FUNCTION_BLOCK Processing2CAT (* CAT Function Block Type *)
  (* Standard: 61499-2 *)
  (* Version 0.0, 7/7/2026, template *)
  PACKAGE Main;
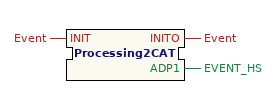
  EVENT_INPUT
    INIT; (* Initialization Request *)
  END_EVENT
  EVENT_OUTPUT
    INITO; (* Initialization Confirm *)
  END_EVENT
  PLUGS
    ADP1 : EVENT_HS;
  END_PLUGS
  FBS
    FB1 : ProcessingSequence1;
    FB2 : TableDriver;
    Tester : SingleActingActuator;
    Drill : DrillDriver;
    FB5 : SYMLINKMULTIVARDST_238520AAD20108C65(QI := TRUE, NAME1 := '$${PATH}WP_AVAIL', NAME2 := '$${PATH}WP_DRILL', NAME3 := '$${PATH}WP_TEST', NAME4 := '$${PATH}DRILL_RAISED', NAME5 := '$${PATH}DRILL_LOWERED', NAME6 := '$${PATH}IN_POSITION', NAME7 := '$${PATH}HOLE_DETECTED'); {SET_ATTRIBUTE(Configuration.GenericFBType.InterfaceParams, Runtime.System#I:=7;VALUE${I$}:BOOL,BOOL,BOOL,BOOL,BOOL,BOOL,BOOL)}
    FB7 : SYMLINKMULTIVARSRC_5495E501E675F500(QI := TRUE, NAME1 := '$${PATH}START_DRILL', NAME2 := '$${PATH}ROTATE', NAME3 := '$${PATH}LOWER_DRILL', NAME4 := '$${PATH}RAISE_DRILL', NAME5 := '$${PATH}CLAMP', NAME6 := '$${PATH}TEST'); {SET_ATTRIBUTE(Configuration.GenericFBType.InterfaceParams, Runtime.System#I:=6;VALUE${I$}:BOOL,BOOL,BOOL,BOOL,BOOL,BOOL)}
    Clamp : SingleActingActuator;
  END_FBS
  EVENT_CONNECTIONS
    ADP1.06D0DEC05BDF54B5 TO FB1.C97AC495352E3E1E;
    FB1.B088E5234850CB03 TO ADP1.17D55D3741201415;
    INIT TO FB5.INIT;
    FB1.D3B5A8B772FCEA74 TO FB2.6DA377513BB052A8;
    FB1.0CDBBA126F3EB67D TO FB2.BE47842DE556BB00;
    FB1.C353476483DC6313 TO Tester.CCF810354971381B;
    FB1.146D4250297CC697 TO Tester.1BF27B5DCFCCFAF4;
    FB1.A987DB2144D107B9 TO Drill.1D30737806201FD6;
    FB1.1FE929CFCAA94308 TO Drill.0BFE808CC7BF5304;
    FB1.F82CF39030B50881 TO Drill.894E27CD5DAB3D2C;
    FB1.0FC9D8B2B29AA22D TO Drill.CDBB9A3D25440EBE;
    FB1.97F5D70C41BD3D18 TO Clamp.1BF27B5DCFCCFAF4;
    FB1.A8BDF88CF1CF6D8D TO Clamp.CCF810354971381B;
    FB5.CNF TO FB1.C1A7677E5176E42B;
    FB5.CNF TO FB2.1CCD0C1482531427;
    FB5.CNF TO Drill.07A841519EEF7D29;
    FB5.INITO TO FB7.INIT;
    Drill.B515F055283B6D1D TO FB7.REQ;
    Clamp.BC8FA2DBFA3F03EE TO FB7.REQ;
    Drill.2184ADB07913F188 TO FB7.REQ;
    Tester.BC8FA2DBFA3F03EE TO FB7.REQ;
    FB2.2F1CB770CB922D4B TO FB7.REQ;
    FB7.INITO TO INITO;
    FB7.INITO TO FB2.C2FC305C6C7872B8;
    FB7.INITO TO Tester.A4B796CDD9024B67;
    FB7.INITO TO Drill.82E100EB26E04504;
    FB7.INITO TO Clamp.A4B796CDD9024B67;
  END_CONNECTIONS
  DATA_CONNECTIONS
    FB5.VALUE2 TO FB1.E1F7FAE400B6E48F;
    FB5.VALUE3 TO FB1.77895791E5012799;
    FB5.VALUE4 TO FB1.909F52C6313386F9;
    FB5.VALUE4 TO Drill.113F4B319C5D4EEB;
    FB5.VALUE5 TO FB1.93B5E068BF203B9B;
    FB5.VALUE5 TO Drill.FC5030D73ADCE20B;
    FB5.VALUE6 TO FB1.D00EBC763795CCDE;
    FB5.VALUE6 TO FB2.B3C88798EBFDA44D;
    FB5.VALUE7 TO FB1.91161A4E26D35ED7;
    Drill.137A4746C9FE30DB TO FB7.VALUE1;
    FB2.E31FA5EA69A50141 TO FB7.VALUE2;
    Drill.1A5F06F8AAA23A4B TO FB7.VALUE3;
    Drill.349DADD9FC043770 TO FB7.VALUE4;
    Clamp.74B9BF94DC489173 TO FB7.VALUE5;
    Tester.74B9BF94DC489173 TO FB7.VALUE6;
  END_CONNECTIONS
END_FUNCTION_BLOCK
